FUNCTION_BLOCK ARM_CONTROL
  {SET_ATTRIBUTE(OpcUa, SERVICE)}
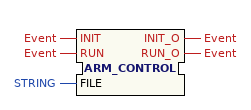
  EVENT_INPUT
    INIT;
    RUN;
  END_EVENT
  EVENT_OUTPUT
    INIT_O;
    RUN_O;
  END_EVENT
  VAR_INPUT
    FILE : STRING;
  END_VAR
END_FUNCTION_BLOCK
